{attribute 'qualified_only'}
VAR_GLOBAL
    stLivingRoomCeilingCmd : ST_LightCmd;
    stLivingRoomWallCmd    : ST_LightCmd;
    stLivingRoomAmbientCmd : ST_LightCmd;
END_VAR

(* stored: Version 1.1.0.1, ProductVersion 3.1.4026.20
   GVL GVL_LightCmds: Id {A8100003-3B71-4C96-8F25-7A1B2C3D4001} *)
